(* IEC 61131-3 sources: llm-plc-st-eval/codesys/_respaldo_20260909, 9 files *)

(* ---- PRG_Test_B4.st ---- *)
(*) Banco B4. violacionInterlock se muestrea y enclava en CADA scan. *)
PROGRAM PRG_Test_B4
VAR CONSTANT ULTIMO_PASO : INT := 7; END_VAR
VAR
 fb: FB_Giro; btnFwd,btnRev,btnParo,espFwd,espRev,pulsoReset,finalizado,violacionInterlock: BOOL;
 paso,i,nPasan: INT; tPaso: TON; resultado: ARRAY[0..7] OF INT; veredicto: INT;
END_VAR
tPaso(IN:=NOT pulsoReset,PT:=T#150MS); pulsoReset:=FALSE;
IF NOT finalizado THEN CASE paso OF
 0: btnFwd:=FALSE;btnRev:=FALSE;btnParo:=FALSE;espFwd:=FALSE;espRev:=FALSE; (* reposo *)
 1: btnFwd:=TRUE;espFwd:=TRUE;espRev:=FALSE; (* marcha adelante *)
 2: btnFwd:=FALSE;espFwd:=TRUE;espRev:=FALSE; (* enclavamiento FWD *)
 3: btnRev:=TRUE;espFwd:=TRUE;espRev:=FALSE; (* Rev sin paro: prohibido *)
 4: btnRev:=FALSE;btnParo:=TRUE;espFwd:=FALSE;espRev:=FALSE; (* paro *)
 5: btnParo:=FALSE;btnRev:=TRUE;espFwd:=FALSE;espRev:=TRUE; (* marcha reversa *)
 6: btnFwd:=TRUE;btnRev:=TRUE;espFwd:=FALSE;espRev:=TRUE; (* ambas ordenes: nunca ambas salidas *)
 7: btnFwd:=FALSE;btnRev:=FALSE;btnParo:=TRUE;espFwd:=FALSE;espRev:=FALSE; (* paro final *)
 END_CASE END_IF
fb(btnFwd:=btnFwd,btnRev:=btnRev,btnParo:=btnParo);
IF fb.fwd AND fb.rev THEN violacionInterlock:=TRUE; END_IF;
IF tPaso.Q AND NOT finalizado THEN IF (fb.fwd=espFwd) AND (fb.rev=espRev) THEN resultado[paso]:=1; ELSE resultado[paso]:=2; END_IF; pulsoReset:=TRUE; IF paso<ULTIMO_PASO THEN paso:=paso+1; ELSE finalizado:=TRUE; END_IF END_IF
IF finalizado AND veredicto=0 THEN nPasan:=0;FOR i:=0 TO ULTIMO_PASO DO IF resultado[i]=1 THEN nPasan:=nPasan+1;END_IF END_FOR;IF nPasan=ULTIMO_PASO+1 AND NOT violacionInterlock THEN veredicto:=1;ELSE veredicto:=2;END_IF END_IF

(* ---- PRG_Test_B5.st ---- *)
(*) Banco B5: prueba TOF, tiempo de 30 s y rearme durante post-enfriamiento. *)
PROGRAM PRG_Test_B5
VAR CONSTANT ULTIMO_PASO:INT:=6; END_VAR
VAR fb:FB_Ventilador; quemadorOn,esperado,pulsoReset,finalizado:BOOL;paso,i,nPasan:INT;tEspera:TIME;tPaso:TON;resultado:ARRAY[0..6] OF INT;veredicto:INT;END_VAR
IF NOT finalizado THEN CASE paso OF
0:quemadorOn:=FALSE;tEspera:=T#200MS;esperado:=FALSE;
1:quemadorOn:=TRUE;tEspera:=T#200MS;esperado:=TRUE; (* acompana quemador *)
2:quemadorOn:=FALSE;tEspera:=T#29S;esperado:=TRUE; (* antes de 30 s *)
3:quemadorOn:=FALSE;tEspera:=T#1200MS;esperado:=FALSE; (* 30.2 s acumulados *)
4:quemadorOn:=TRUE;tEspera:=T#200MS;esperado:=TRUE;
5:quemadorOn:=FALSE;tEspera:=T#10S;esperado:=TRUE; (* post-enfriamiento, se reenciende *)
6:quemadorOn:=TRUE;tEspera:=T#200MS;esperado:=TRUE; (* reactivacion reinicia TOF *)
END_CASE END_IF
tPaso(IN:=NOT pulsoReset,PT:=tEspera);pulsoReset:=FALSE;fb(quemadorOn:=quemadorOn);
IF tPaso.Q AND NOT finalizado THEN IF fb.ventilador=esperado THEN resultado[paso]:=1;ELSE resultado[paso]:=2;END_IF;pulsoReset:=TRUE;IF paso<ULTIMO_PASO THEN paso:=paso+1;ELSE finalizado:=TRUE;END_IF END_IF
IF finalizado AND veredicto=0 THEN nPasan:=0;FOR i:=0 TO ULTIMO_PASO DO IF resultado[i]=1 THEN nPasan:=nPasan+1;END_IF END_FOR;IF nPasan=ULTIMO_PASO+1 THEN veredicto:=1;ELSE veredicto:=2;END_IF END_IF

(* ---- PRG_Test_B6.st ---- *)
(*) B6: mide intervalos completos ON/OFF, T#1S +/- T#150MS. MainTask: 4..10 ms. *)
PROGRAM PRG_Test_B6
VAR CONSTANT ULTIMO_PASO:INT:=2;END_VAR
VAR fb:FB_Baliza;alarma,pulsoReset,resetIntervalo,finalizado,prev,primer,error:BOOL;paso,i,nPasan,nOn,nOff:INT;tEspera:TIME;tPaso,tIntervalo:TON;resultado:ARRAY[0..2] OF INT;veredicto:INT;duracion:TIME;END_VAR
IF NOT finalizado THEN CASE paso OF 0:alarma:=FALSE;tEspera:=T#200MS;1:alarma:=TRUE;tEspera:=T#7S;2:alarma:=FALSE;tEspera:=T#200MS;END_CASE END_IF
tPaso(IN:=NOT pulsoReset,PT:=tEspera);tIntervalo(IN:=NOT resetIntervalo,PT:=T#10S);pulsoReset:=FALSE;resetIntervalo:=FALSE;fb(alarma:=alarma);
IF paso=1 THEN
 IF (fb.lampara AND NOT prev) OR ((NOT fb.lampara) AND prev) THEN
  IF primer THEN duracion:=tIntervalo.ET;IF NOT fb.lampara THEN nOn:=nOn+1;ELSE nOff:=nOff+1;END_IF;IF duracion<T#850MS OR duracion>T#1150MS THEN error:=TRUE;END_IF;ELSE primer:=TRUE;END_IF;
  resetIntervalo:=TRUE;
 END_IF
END_IF;prev:=fb.lampara;
IF tPaso.Q AND NOT finalizado THEN
 IF (paso=0 AND NOT fb.lampara) OR (paso=1 AND nOn>=2 AND nOff>=2 AND NOT error) OR (paso=2 AND NOT fb.lampara) THEN resultado[paso]:=1;ELSE resultado[paso]:=2;END_IF;
 pulsoReset:=TRUE;IF paso<ULTIMO_PASO THEN paso:=paso+1;ELSE finalizado:=TRUE;END_IF
END_IF
IF finalizado AND veredicto=0 THEN nPasan:=0;FOR i:=0 TO ULTIMO_PASO DO IF resultado[i]=1 THEN nPasan:=nPasan+1;END_IF END_FOR;IF nPasan=ULTIMO_PASO+1 THEN veredicto:=1;ELSE veredicto:=2;END_IF END_IF

(* ---- PRG_Test_I1.st ---- *)
(*) I1: secuencia 20/4/15 s y amarillo intermitente medido por flancos. *)
PROGRAM PRG_Test_I1
VAR CONSTANT ULTIMO_PASO:INT:=6;END_VAR
VAR fb:FB_Semaforo;habilitado,pulsoReset,resetIntervalo,finalizado,prevA,primer,error,espV,espA,espR:BOOL;paso,i,nPasan,nOn,nOff:INT;tEspera,duracion:TIME;tPaso,tIntervalo:TON;resultado:ARRAY[0..6] OF INT;veredicto:INT;END_VAR
IF NOT finalizado THEN CASE paso OF
0:habilitado:=FALSE;tEspera:=T#200MS;espV:=FALSE;espR:=FALSE;
1:habilitado:=TRUE;tEspera:=T#200MS;espV:=TRUE;espA:=FALSE;espR:=FALSE;
2:habilitado:=TRUE;tEspera:=T#20S;espV:=FALSE;espA:=TRUE;espR:=FALSE;
3:habilitado:=TRUE;tEspera:=T#4S;espV:=FALSE;espA:=FALSE;espR:=TRUE;
4:habilitado:=TRUE;tEspera:=T#15S;espV:=TRUE;espA:=FALSE;espR:=FALSE;
5:habilitado:=FALSE;tEspera:=T#7S;espV:=FALSE;espR:=FALSE;
6:habilitado:=TRUE;tEspera:=T#200MS;espV:=TRUE;espA:=FALSE;espR:=FALSE;END_CASE END_IF
tPaso(IN:=NOT pulsoReset,PT:=tEspera);tIntervalo(IN:=NOT resetIntervalo,PT:=T#10S);pulsoReset:=FALSE;resetIntervalo:=FALSE;fb(habilitado:=habilitado);
IF paso=5 AND ((fb.luzA AND NOT prevA) OR ((NOT fb.luzA) AND prevA)) THEN IF primer THEN duracion:=tIntervalo.ET;IF NOT fb.luzA THEN nOn:=nOn+1;ELSE nOff:=nOff+1;END_IF;IF duracion<T#850MS OR duracion>T#1150MS THEN error:=TRUE;END_IF;ELSE primer:=TRUE;END_IF;resetIntervalo:=TRUE;END_IF;prevA:=fb.luzA;
IF tPaso.Q AND NOT finalizado THEN IF ((paso=0 AND NOT fb.luzV AND NOT fb.luzR) OR (paso>=1 AND paso<>5 AND fb.luzV=espV AND fb.luzA=espA AND fb.luzR=espR) OR (paso=5 AND NOT fb.luzV AND NOT fb.luzR AND nOn>=2 AND nOff>=2 AND NOT error)) THEN resultado[paso]:=1;ELSE resultado[paso]:=2;END_IF;pulsoReset:=TRUE;IF paso<ULTIMO_PASO THEN paso:=paso+1;ELSE finalizado:=TRUE;END_IF END_IF
IF finalizado AND veredicto=0 THEN nPasan:=0;FOR i:=0 TO ULTIMO_PASO DO IF resultado[i]=1 THEN nPasan:=nPasan+1;END_IF END_FOR;IF nPasan=ULTIMO_PASO+1 THEN veredicto:=1;ELSE veredicto:=2;END_IF END_IF

(* ---- PRG_Test_I2.st ---- *)
(*) I2: orden de estados, temporizacion de mezcla y paro seguro en dos fases. *)
PROGRAM PRG_Test_I2
VAR CONSTANT ULTIMO_PASO:INT:=9;END_VAR
VAR fb:FB_Llenado;nivelAlto,nivelBajo,btnInicio,btnParo,evL,evM,evD,pulsoReset,finalizado:BOOL;paso,i,nPasan:INT;tEspera:TIME;tPaso:TON;resultado:ARRAY[0..9] OF INT;veredicto:INT;END_VAR
IF NOT finalizado THEN CASE paso OF
0:nivelAlto:=FALSE;nivelBajo:=FALSE;btnInicio:=FALSE;btnParo:=FALSE;tEspera:=T#200MS;evL:=FALSE;evM:=FALSE;evD:=FALSE;
1:btnInicio:=TRUE;tEspera:=T#200MS;evL:=TRUE;evM:=FALSE;evD:=FALSE;
2:btnInicio:=FALSE;nivelAlto:=TRUE;tEspera:=T#200MS;evL:=FALSE;evM:=TRUE;evD:=FALSE;
3:tEspera:=T#59800MS;evM:=TRUE; (* antes de 60 s *)
4:tEspera:=T#500MS;evL:=FALSE;evM:=FALSE;evD:=TRUE;
5:nivelBajo:=TRUE;tEspera:=T#200MS;evL:=FALSE;evM:=FALSE;evD:=FALSE;
6:nivelAlto:=FALSE;nivelBajo:=FALSE;btnInicio:=TRUE;tEspera:=T#200MS;evL:=TRUE;evM:=FALSE;evD:=FALSE;
7:btnInicio:=FALSE;btnParo:=TRUE;tEspera:=T#200MS;evL:=FALSE;evM:=FALSE;evD:=FALSE; (* paro en llenado *)
8:btnParo:=FALSE;btnInicio:=TRUE;tEspera:=T#200MS;evL:=TRUE;evM:=FALSE;evD:=FALSE;
9:btnInicio:=FALSE;nivelAlto:=TRUE;btnParo:=TRUE;tEspera:=T#200MS;evL:=FALSE;evM:=FALSE;evD:=FALSE; (* paro en mezcla *) END_CASE END_IF
tPaso(IN:=NOT pulsoReset,PT:=tEspera);pulsoReset:=FALSE;fb(nivelAlto:=nivelAlto,nivelBajo:=nivelBajo,btnInicio:=btnInicio,btnParo:=btnParo);
IF tPaso.Q AND NOT finalizado THEN IF fb.vLlenado=evL AND fb.motorMezcla=evM AND fb.vDescarga=evD THEN resultado[paso]:=1;ELSE resultado[paso]:=2;END_IF;pulsoReset:=TRUE;IF paso<ULTIMO_PASO THEN paso:=paso+1;ELSE finalizado:=TRUE;END_IF END_IF
IF finalizado AND veredicto=0 THEN nPasan:=0;FOR i:=0 TO ULTIMO_PASO DO IF resultado[i]=1 THEN nPasan:=nPasan+1;END_IF END_FOR;IF nPasan=ULTIMO_PASO+1 THEN veredicto:=1;ELSE veredicto:=2;END_IF END_IF

(* ---- PRG_Test_I3.st ---- *)
(*) Banco I3: retencion individual, ACK condicionado y prioridad. *)
PROGRAM PRG_Test_I3
VAR CONSTANT ULTIMO_PASO:INT:=8;END_VAR
VAR fb:FB_Alarmas;alm1,alm2,alm3,ack1,ack2,ack3,espSirena,pulsoReset,finalizado:BOOL;espCodigo,paso,i,nPasan:INT;tPaso:TON;resultado:ARRAY[0..8] OF INT;veredicto:INT;END_VAR
tPaso(IN:=NOT pulsoReset,PT:=T#150MS);pulsoReset:=FALSE;
IF NOT finalizado THEN CASE paso OF
0:alm1:=FALSE;alm2:=FALSE;alm3:=FALSE;ack1:=TRUE;ack2:=TRUE;ack3:=TRUE;espSirena:=FALSE;espCodigo:=0;
1:ack1:=FALSE;ack2:=FALSE;ack3:=FALSE;alm3:=TRUE;espSirena:=TRUE;espCodigo:=3;
2:alm3:=FALSE;espSirena:=TRUE;espCodigo:=3; (* retencion *)
3:ack3:=TRUE;espSirena:=FALSE;espCodigo:=0; (* ACK al retirar causa *)
4:ack3:=FALSE;alm2:=TRUE;alm3:=TRUE;espSirena:=TRUE;espCodigo:=2;
5:alm1:=TRUE;espSirena:=TRUE;espCodigo:=1; (* prioridad alta *)
6:alm1:=FALSE;ack1:=TRUE;espSirena:=TRUE;espCodigo:=2;
7:alm2:=FALSE;ack2:=TRUE;espSirena:=TRUE;espCodigo:=3;
8:alm3:=FALSE;ack3:=TRUE;espSirena:=FALSE;espCodigo:=0;
END_CASE END_IF
fb(alm1:=alm1,alm2:=alm2,alm3:=alm3,ack1:=ack1,ack2:=ack2,ack3:=ack3);
IF tPaso.Q AND NOT finalizado THEN IF fb.sirena=espSirena AND fb.codigoAlm=espCodigo THEN resultado[paso]:=1;ELSE resultado[paso]:=2;END_IF;pulsoReset:=TRUE;IF paso<ULTIMO_PASO THEN paso:=paso+1;ELSE finalizado:=TRUE;END_IF END_IF
IF finalizado AND veredicto=0 THEN nPasan:=0;FOR i:=0 TO ULTIMO_PASO DO IF resultado[i]=1 THEN nPasan:=nPasan+1;END_IF END_FOR;IF nPasan=ULTIMO_PASO+1 THEN veredicto:=1;ELSE veredicto:=2;END_IF END_IF

(* ---- PRG_Test_I4.st ---- *)
(*) I4: interlock enclavado y tiempo muerto medido entre caida kY y subida kD. MainTask 4..10 ms. *)
PROGRAM PRG_Test_I4
VAR CONSTANT ULTIMO_PASO:INT:=5;END_VAR
VAR fb:FB_EstrellaTriangulo;btnMarcha,btnParo,pulsoReset,resetMed,finalizado,prevY,prevD,midiendo,interlock,muertoOK:BOOL;paso,i,nPasan:INT;tEspera,duracionMuerto:TIME;tPaso,tMed:TON;resultado:ARRAY[0..5] OF INT;veredicto:INT;END_VAR
IF NOT finalizado THEN CASE paso OF 0:btnMarcha:=FALSE;btnParo:=FALSE;tEspera:=T#200MS;1:btnMarcha:=TRUE;tEspera:=T#7800MS;2:btnMarcha:=TRUE;tEspera:=T#500MS;3:btnMarcha:=TRUE;tEspera:=T#300MS;4:btnMarcha:=FALSE;btnParo:=TRUE;tEspera:=T#200MS;5:btnParo:=FALSE;btnMarcha:=TRUE;tEspera:=T#200MS;END_CASE END_IF
tPaso(IN:=NOT pulsoReset,PT:=tEspera);tMed(IN:=NOT resetMed,PT:=T#10S);pulsoReset:=FALSE;resetMed:=FALSE;fb(btnMarcha:=btnMarcha,btnParo:=btnParo);
IF fb.kY AND fb.kD THEN interlock:=TRUE;END_IF;
IF prevY AND NOT fb.kY THEN midiendo:=TRUE;resetMed:=TRUE;END_IF;
IF midiendo AND fb.kD AND NOT prevD THEN duracionMuerto:=tMed.ET;IF duracionMuerto>=T#100MS THEN muertoOK:=TRUE;END_IF;midiendo:=FALSE;END_IF;prevY:=fb.kY;prevD:=fb.kD;
IF tPaso.Q AND NOT finalizado THEN IF (paso=0 AND NOT fb.kM AND NOT fb.kY AND NOT fb.kD) OR (paso=1 AND fb.kM AND fb.kY AND NOT fb.kD) OR (paso=2 AND fb.kM AND NOT fb.kY AND NOT fb.kD) OR (paso=3 AND fb.kM AND NOT fb.kY AND fb.kD AND muertoOK) OR (paso=4 AND NOT fb.kM AND NOT fb.kY AND NOT fb.kD) OR (paso=5 AND fb.kM AND fb.kY AND NOT fb.kD) THEN resultado[paso]:=1;ELSE resultado[paso]:=2;END_IF;pulsoReset:=TRUE;IF paso<ULTIMO_PASO THEN paso:=paso+1;ELSE finalizado:=TRUE;END_IF END_IF
IF finalizado AND veredicto=0 THEN nPasan:=0;FOR i:=0 TO ULTIMO_PASO DO IF resultado[i]=1 THEN nPasan:=nPasan+1;END_IF END_FOR;IF nPasan=ULTIMO_PASO+1 AND NOT interlock THEN veredicto:=1;ELSE veredicto:=2;END_IF END_IF

(* ---- PRG_Test_I5.st ---- *)
(*) I5: presencia sostenida no puede contar mas de una pieza; desvio 2 s + 1 s. *)
PROGRAM PRG_Test_I5
VAR CONSTANT ULTIMO_PASO:INT:=6;END_VAR
VAR fb:FB_Clasificadora;sensorPresencia,sensorAltura,pulsoReset,finalizado,espBanda,espPiston:BOOL;espAltas,espBajas,paso,i,nPasan:INT;tEspera:TIME;tPaso:TON;resultado:ARRAY[0..6] OF INT;veredicto:INT;END_VAR
IF NOT finalizado THEN CASE paso OF
0:sensorPresencia:=FALSE;sensorAltura:=FALSE;tEspera:=T#200MS;espBanda:=TRUE;espPiston:=FALSE;espAltas:=0;espBajas:=0;
1:sensorPresencia:=TRUE;sensorAltura:=FALSE;tEspera:=T#300MS;espBanda:=TRUE;espPiston:=FALSE;espAltas:=0;espBajas:=1; (* baja sostenida *)
2:sensorPresencia:=FALSE;tEspera:=T#200MS;espBanda:=TRUE;espPiston:=FALSE;espAltas:=0;espBajas:=1;
3:sensorPresencia:=TRUE;sensorAltura:=TRUE;tEspera:=T#200MS;espBanda:=TRUE;espPiston:=FALSE;espAltas:=1;espBajas:=1;
4:sensorPresencia:=FALSE;sensorAltura:=FALSE;tEspera:=T#1800MS;espBanda:=TRUE;espPiston:=FALSE;espAltas:=1;espBajas:=1; (* antes de 2 s *)
5:tEspera:=T#400MS;espBanda:=TRUE;espPiston:=TRUE;espAltas:=1;espBajas:=1; (* dentro del pulso *)
6:tEspera:=T#1200MS;espBanda:=TRUE;espPiston:=FALSE;espAltas:=1;espBajas:=1;END_CASE END_IF
tPaso(IN:=NOT pulsoReset,PT:=tEspera);pulsoReset:=FALSE;fb(sensorPresencia:=sensorPresencia,sensorAltura:=sensorAltura);
IF tPaso.Q AND NOT finalizado THEN IF fb.banda=espBanda AND fb.piston=espPiston AND fb.nAltas=espAltas AND fb.nBajas=espBajas THEN resultado[paso]:=1;ELSE resultado[paso]:=2;END_IF;pulsoReset:=TRUE;IF paso<ULTIMO_PASO THEN paso:=paso+1;ELSE finalizado:=TRUE;END_IF END_IF
IF finalizado AND veredicto=0 THEN nPasan:=0;FOR i:=0 TO ULTIMO_PASO DO IF resultado[i]=1 THEN nPasan:=nPasan+1;END_IF END_FOR;IF nPasan=ULTIMO_PASO+1 THEN veredicto:=1;ELSE veredicto:=2;END_IF END_IF

(* ---- PRG_Test_I6.st ---- *)
(*) I6: escalado 0..27648 a 0..100 y ambos sentidos de la histéresis. *)
PROGRAM PRG_Test_I6
VAR CONSTANT ULTIMO_PASO:INT:=7;END_VAR
VAR fb:FB_Temperatura;rawTemp,espRaw,paso,i,nPasan:INT;espTemp:REAL;espFrio,espAlarma,pulsoReset,finalizado:BOOL;tPaso:TON;resultado:ARRAY[0..7] OF INT;veredicto:INT;END_VAR
tPaso(IN:=NOT pulsoReset,PT:=T#100MS);pulsoReset:=FALSE;
IF NOT finalizado THEN CASE paso OF
0:rawTemp:=13824;espTemp:=50.0;espFrio:=FALSE;espAlarma:=FALSE;
1:rawTemp:=22119;espTemp:=80.0;espFrio:=TRUE;espAlarma:=FALSE;
2:rawTemp:=21289;espTemp:=77.0;espFrio:=TRUE;espAlarma:=FALSE; (* banda: conserva ON *)
3:rawTemp:=20736;espTemp:=75.0;espFrio:=FALSE;espAlarma:=FALSE;
4:rawTemp:=21289;espTemp:=77.0;espFrio:=FALSE;espAlarma:=FALSE; (* banda: conserva OFF *)
5:rawTemp:=27649;espTemp:=0.0;espFrio:=FALSE;espAlarma:=TRUE;
6:rawTemp:=-1;espTemp:=0.0;espFrio:=FALSE;espAlarma:=TRUE;
7:rawTemp:=0;espTemp:=0.0;espFrio:=FALSE;espAlarma:=FALSE;END_CASE END_IF
fb(rawTemp:=rawTemp);
IF tPaso.Q AND NOT finalizado THEN IF ((paso>=5) OR ((fb.tempC>espTemp-0.1) AND (fb.tempC<espTemp+0.1))) AND fb.enfriador=espFrio AND fb.almSensor=espAlarma THEN resultado[paso]:=1;ELSE resultado[paso]:=2;END_IF;pulsoReset:=TRUE;IF paso<ULTIMO_PASO THEN paso:=paso+1;ELSE finalizado:=TRUE;END_IF END_IF
IF finalizado AND veredicto=0 THEN nPasan:=0;FOR i:=0 TO ULTIMO_PASO DO IF resultado[i]=1 THEN nPasan:=nPasan+1;END_IF END_FOR;IF nPasan=ULTIMO_PASO+1 THEN veredicto:=1;ELSE veredicto:=2;END_IF END_IF
